Fanuc KAREL source: ka00118.KL

-- PROVISIONAL review KL for V940-1; original PC SHA256 f4b33f0ee74c0066efe5c3a563572c282fd395e2a2b907961120658c159d31c7
-- Incomplete behavior may be omitted. Consult companion uncertainty JSON. Do not deploy.
PROGRAM KA00118
%NOLOCKGROUP
-- UNRESOLVED_DECL SRC type=00001c
-- UNRESOLVED_DECL DST type=00001c
BEGIN
  -- V9_ZERO_TABLE_METADATA_HINT layout=0001; no indexed target words; source/name/runtime held
  -- UNRESOLVED_PC offsets 5-15; opcodes 9D,22,A5
  -- UNRESOLVED_PC offsets 20-32; opcodes 21,23
  -- UNRESOLVED_PC offsets 37-41; opcodes 7F
END KA00118
